Fanuc KAREL source: kt00040.KL

-- PROVISIONAL review KL for V770-1; original PC SHA256 79837d10b995025f10d2a3231018bcf29c137b4d7d4045e5310f95cecba7086b
-- Incomplete behavior may be omitted. Consult companion uncertainty JSON. Do not deploy.
PROGRAM KT00040
%NOLOCKGROUP
VAR
  I1 : INTEGER
  OUT : REAL
-- UNRESOLVED_DECL H2 type=002017
BEGIN
  -- UNRESOLVED_PC offsets 5-16; opcodes 2E,23
  -- UNRESOLVED_PC offsets 21-35; opcodes 2E,22,9D,33,B4
  -- UNRESOLVED_PC offsets 40-63; opcodes 21,22,9D,33,B3,53,64,23
  -- UNRESOLVED_PC offsets 68-72; opcodes 7F
END KT00040
